FUNCTION_BLOCK BATCH_FILLING (* Migrated from IEC 61131-3 ST *)
  (* Standard: 61499-2 *)
  (* Version 1.0, 2026-11-06, st2fb *)
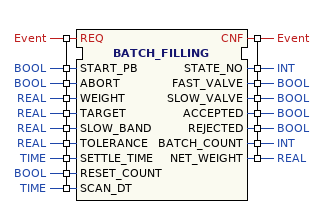
  EVENT_INPUT
    REQ WITH START_PB, ABORT, WEIGHT, TARGET, SLOW_BAND, TOLERANCE, SETTLE_TIME, RESET_COUNT, SCAN_DT;
  END_EVENT
  EVENT_OUTPUT
    CNF WITH STATE_NO, FAST_VALVE, SLOW_VALVE, ACCEPTED, REJECTED, BATCH_COUNT, NET_WEIGHT;
  END_EVENT
  VAR_INPUT
    START_PB : BOOL;
    ABORT : BOOL;
    WEIGHT : REAL;
    TARGET : REAL;
    SLOW_BAND : REAL;
    TOLERANCE : REAL;
    SETTLE_TIME : TIME;
    RESET_COUNT : BOOL;
    SCAN_DT : TIME;
  END_VAR
  VAR_OUTPUT
    STATE_NO : INT;
    FAST_VALVE : BOOL;
    SLOW_VALVE : BOOL;
    ACCEPTED : BOOL;
    REJECTED : BOOL;
    BATCH_COUNT : INT;
    NET_WEIGHT : REAL;
  END_VAR
  VAR
    TARE : REAL := 0.0;
    COUNT_PULSE : BOOL := FALSE;
    ST2FB_NOW : TIME := T#0s;
    START_EDGE_CLK : BOOL := FALSE;
    START_EDGE_Q : BOOL := FALSE;
    START_EDGE_M : BOOL := FALSE;
    SETTLE_TIMER_IN : BOOL := FALSE;
    SETTLE_TIMER_PT : TIME := T#0s;
    SETTLE_TIMER_Q : BOOL := FALSE;
    SETTLE_TIMER_ET : TIME := T#0s;
    SETTLE_TIMER_STATE : INT := 0;
    SETTLE_TIMER_PREV_IN : BOOL := FALSE;
    SETTLE_TIMER_START_TIME : TIME := T#0s;
    COUNTER_CU : BOOL := FALSE;
    COUNTER_R : BOOL := FALSE;
    COUNTER_PV : INT := 0;
    COUNTER_Q : BOOL := FALSE;
    COUNTER_CV : INT := 0;
    COUNTER_CU_T_Q : BOOL := FALSE;
    COUNTER_CU_T_M : BOOL := FALSE;
  END_VAR
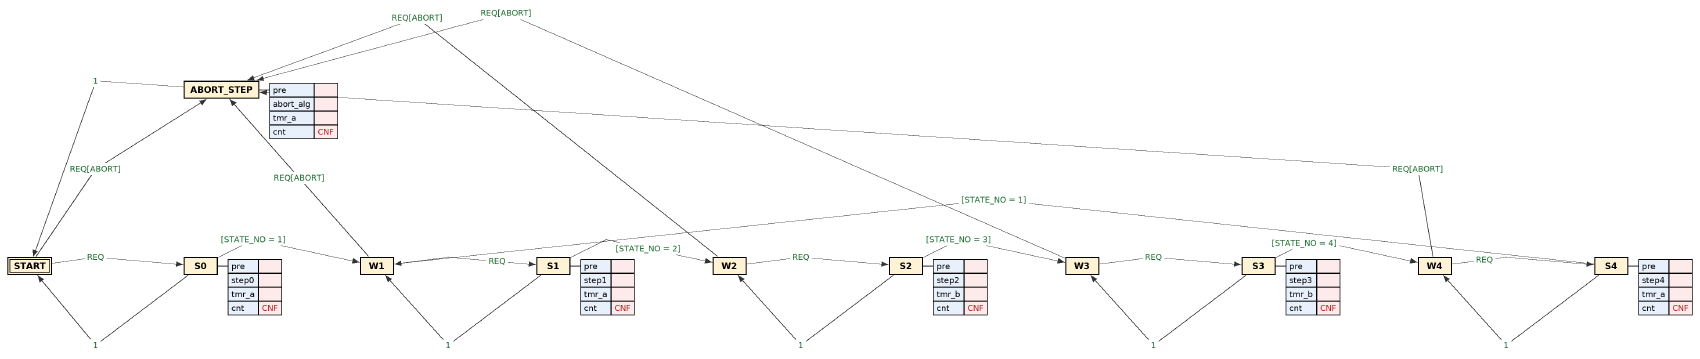
  EC_STATES
    START;
    ABORT_STEP : pre, abort_alg, tmr_a, cnt -> CNF;
    S0 : pre, step0, tmr_a, cnt -> CNF;
    W1;
    S1 : pre, step1, tmr_a, cnt -> CNF;
    W2;
    S2 : pre, step2, tmr_b, cnt -> CNF;
    W3;
    S3 : pre, step3, tmr_b, cnt -> CNF;
    W4;
    S4 : pre, step4, tmr_a, cnt -> CNF;
  END_STATES
  EC_TRANSITIONS
    START TO ABORT_STEP := REQ[ABORT];
    START TO S0 := REQ;
    ABORT_STEP TO START := 1;
    S0 TO W1 := [STATE_NO = 1];
    S0 TO START := 1;
    W1 TO ABORT_STEP := REQ[ABORT];
    W1 TO S1 := REQ;
    S1 TO W2 := [STATE_NO = 2];
    S1 TO W1 := 1;
    W2 TO ABORT_STEP := REQ[ABORT];
    W2 TO S2 := REQ;
    S2 TO W3 := [STATE_NO = 3];
    S2 TO W2 := 1;
    W3 TO ABORT_STEP := REQ[ABORT];
    W3 TO S3 := REQ;
    S3 TO W4 := [STATE_NO = 4];
    S3 TO W3 := 1;
    W4 TO ABORT_STEP := REQ[ABORT];
    W4 TO S4 := REQ;
    S4 TO W1 := [STATE_NO = 1];
    S4 TO W4 := 1;
  END_TRANSITIONS
  ALGORITHM pre IN ST:
ST2FB_NOW := ST2FB_NOW + SCAN_DT;
START_EDGE_CLK := START_PB;
START_EDGE_Q := START_EDGE_CLK AND NOT START_EDGE_M;
START_EDGE_M := START_EDGE_CLK;
NET_WEIGHT := WEIGHT - TARE;
FAST_VALVE := FALSE;
SLOW_VALVE := FALSE;
COUNT_PULSE := FALSE;
  END_ALGORITHM
  ALGORITHM abort_alg IN ST:
STATE_NO := 0;
ACCEPTED := FALSE;
REJECTED := FALSE;
  END_ALGORITHM
  ALGORITHM step0 IN ST:
IF START_EDGE_Q AND NOT ABORT THEN
  TARE := WEIGHT;
  NET_WEIGHT := 0.0;
  ACCEPTED := FALSE;
  REJECTED := FALSE;
  STATE_NO := 1;
END_IF;
  END_ALGORITHM
  ALGORITHM step1 IN ST:
FAST_VALVE := TRUE;
SLOW_VALVE := TRUE;
IF NET_WEIGHT >= TARGET - SLOW_BAND THEN
  STATE_NO := 2;
END_IF;
  END_ALGORITHM
  ALGORITHM step2 IN ST:
SLOW_VALVE := TRUE;
IF NET_WEIGHT >= TARGET THEN
  STATE_NO := 3;
END_IF;
  END_ALGORITHM
  ALGORITHM step3 IN ST:
IF SETTLE_TIMER_Q THEN
  IF (NET_WEIGHT >= TARGET - TOLERANCE) AND (NET_WEIGHT <= TARGET + TOLERANCE) THEN
    ACCEPTED := TRUE;
    COUNT_PULSE := TRUE;
  ELSE
    REJECTED := TRUE;
  END_IF;
  STATE_NO := 4;
END_IF;
  END_ALGORITHM
  ALGORITHM step4 IN ST:
IF START_EDGE_Q THEN
  TARE := WEIGHT;
  NET_WEIGHT := 0.0;
  ACCEPTED := FALSE;
  REJECTED := FALSE;
  STATE_NO := 1;
END_IF;
  END_ALGORITHM
  ALGORITHM tmr_a IN ST:
SETTLE_TIMER_IN := FALSE;
SETTLE_TIMER_PT := SETTLE_TIME;
IF (SETTLE_TIMER_STATE = 0) AND NOT SETTLE_TIMER_PREV_IN AND SETTLE_TIMER_IN THEN
  SETTLE_TIMER_STATE := 1;
  SETTLE_TIMER_Q := FALSE;
  SETTLE_TIMER_START_TIME := ST2FB_NOW;
ELSE
  IF NOT SETTLE_TIMER_IN THEN
    SETTLE_TIMER_ET := T#0s;
    SETTLE_TIMER_Q := FALSE;
    SETTLE_TIMER_STATE := 0;
  ELSIF SETTLE_TIMER_STATE = 1 THEN
    IF SETTLE_TIMER_START_TIME + SETTLE_TIMER_PT <= ST2FB_NOW THEN
      SETTLE_TIMER_STATE := 2;
      SETTLE_TIMER_Q := TRUE;
      SETTLE_TIMER_ET := SETTLE_TIMER_PT;
    ELSE
      SETTLE_TIMER_ET := ST2FB_NOW - SETTLE_TIMER_START_TIME;
    END_IF;
  END_IF;
END_IF;
SETTLE_TIMER_PREV_IN := SETTLE_TIMER_IN;
  END_ALGORITHM
  ALGORITHM tmr_b IN ST:
SETTLE_TIMER_IN := (STATE_NO = 3);
SETTLE_TIMER_PT := SETTLE_TIME;
IF (SETTLE_TIMER_STATE = 0) AND NOT SETTLE_TIMER_PREV_IN AND SETTLE_TIMER_IN THEN
  SETTLE_TIMER_STATE := 1;
  SETTLE_TIMER_Q := FALSE;
  SETTLE_TIMER_START_TIME := ST2FB_NOW;
ELSE
  IF NOT SETTLE_TIMER_IN THEN
    SETTLE_TIMER_ET := T#0s;
    SETTLE_TIMER_Q := FALSE;
    SETTLE_TIMER_STATE := 0;
  ELSIF SETTLE_TIMER_STATE = 1 THEN
    IF SETTLE_TIMER_START_TIME + SETTLE_TIMER_PT <= ST2FB_NOW THEN
      SETTLE_TIMER_STATE := 2;
      SETTLE_TIMER_Q := TRUE;
      SETTLE_TIMER_ET := SETTLE_TIMER_PT;
    ELSE
      SETTLE_TIMER_ET := ST2FB_NOW - SETTLE_TIMER_START_TIME;
    END_IF;
  END_IF;
END_IF;
SETTLE_TIMER_PREV_IN := SETTLE_TIMER_IN;
  END_ALGORITHM
  ALGORITHM cnt IN ST:
COUNTER_CU := COUNT_PULSE;
COUNTER_R := RESET_COUNT;
COUNTER_PV := 1000;
COUNTER_CU_T_Q := COUNTER_CU AND NOT COUNTER_CU_T_M;
COUNTER_CU_T_M := COUNTER_CU;
IF COUNTER_R THEN
  COUNTER_CV := 0;
ELSIF COUNTER_CU_T_Q AND (COUNTER_CV < COUNTER_PV) THEN
  COUNTER_CV := COUNTER_CV + 1;
END_IF;
COUNTER_Q := COUNTER_CV >= COUNTER_PV;
BATCH_COUNT := COUNTER_CV;
  END_ALGORITHM
END_FUNCTION_BLOCK
